(* IEC 61131-3 sources: HypervisionPLC-SCADA/demo/varme-plc, 5 files *)

(* ---- globals.st ---- *)
GLOBAL_VAR
  g_cmd    : INT;   (* L1: b0-3 P1-P4, b4 MVS1, b5 MVS2, b6 pille, b7 VP *)
  g_fb     : INT;   (* L2: b0-3 pumpe koerer, b6 pilleflamme, b9 FF-flamme, b10 Laddomat, b11 pillefejl *)
  g_fault  : INT;   (* L4: b0-3 pumpefejl, b4 pille, b5 laekage, b7 VP; b12 VP-fejlsignal *)
  g_speed  : REAL;  (* L4: tidsfaktor *)
  g_tude   : REAL;  (* L4: udetemp *)
  g_att1   : REAL;  (* L3: tank top *)
  g_att3   : REAL;  (* L3: tank midt *)
  g_att6   : REAL;  (* L3: tank bund *)
  g_fftf   : REAL;  (* L2 *)
  g_pftf   : REAL;  (* L2 *)
  g_mch    : REAL;  (* L2: ladeflow til tank kg/s *)
  g_tch    : REAL;  (* L2: ladetemp *)
  g_str    : REAL;  (* L3: vandet til M1 = pillefyrets indloeb (STR eller tanktop) *)
  g_vptf   : REAL;  (* L4: VP-fremloeb til tanken *)
  g_stf_sp : REAL;  (* L1: fremloebssetpunkt *)
  g_tryk   : REAL;  (* L4: bar *)
END_VAR

(* ---- logic1_styring.st ---- *)
PROGRAM Styring
(* Demo-varmeanlaeg, Logic1: styringen (det en rigtig PLC ville goere).
   Laeser anlaeggets tilstand fra GLOBAL_VAR og skriver kommandoer i g_cmd.
   cmd_mode: 0 Auto, 1 Manuel mode 1, 2 Manuel mode 2, 3 Manuel mode 3.
   MODE 1 Hus + pille (M1 AB-A, M2 AB-A, P1) - 2 Hus + pille + tank (M1 AB-A, M2 AB-B, P1)
   - 3 Hus + tank (M1 AB-B, M2 AB-B, P2). Auto: tanken ind (mode 3) ved ATT1 >= sp_tank_ind,
   ud (mode 1) under sp_tank_ud. Varmepumpen startes manuelt (cmd_vp). Interval 500 ms. *)
VAR
  SMS_TXT      : STRING;
  cmd_mode     : INT;
  cmd_kvitter  : BOOL;
  cmd_vp       : BOOL;
  sp_rum       : REAL := 21.0;
  sp_kurve     : REAL := 1.0;
  sp_stf_max   : REAL := 55.0;
  sp_tank_ind  : REAL := 60.0;
  sp_tank_ud   : REAL := 45.0;
  sp_vp_min    : REAL;          (* -5,0 saettes ved foerste scan: negative startvaerdier bliver 0 i firmwaren *)
  MODE         : INT := 1;
  SMS          : INT;
  STF_SP       : REAL;
  TANK_IND     : BOOL;
  PS1          : BOOL;
  PS2          : BOOL;
  PS3          : BOOL;
  PS4          : BOOL;
  F_HUS        : BOOL;
  F_PILLE      : BOOL;
  F_TANK       : BOOL;
  F_BYPASS     : BOOL;
  AL_P1        : BOOL;
  AL_P2        : BOOL;
  AL_P3        : BOOL;
  AL_P4        : BOOL;
  AL_VP        : BOOL;
  AL_PILLE     : BOOL;
  AL_TRYK_LAV  : BOOL;
  AL_TRYK_HOEJ : BOOL;
  AL_FF_TEMP   : BOOL;
  AL_TANK_KOLD : BOOL;
  ALARMER      : INT;
  kv           : BOOL;
  fb           : INT;
  cmd          : INT;
  tude         : REAL;
  t1           : REAL;
  trykstop     : BOOL;
  c_p1         : BOOL;
  c_p2         : BOOL;
  c_p3         : BOOL;
  c_p4         : BOOL;
  c_pille      : BOOL;
  c_vp         : BOOL;
  init         : BOOL;
END_VAR
BEGIN
  IF NOT init THEN sp_vp_min := -5.0; init := TRUE; END_IF;
  kv := cmd_kvitter;
  cmd_kvitter := FALSE;
  fb := g_fb;
  tude := g_tude;
  t1 := g_att1;

  (* Pumpefejl: kommanderet, men ingen tilbagemelding i 10 s -> laast til kvittering *)
  AL_P1 := SR(TON(BIT_TST(g_cmd, 0) AND NOT BIT_TST(fb, 0), T#10s), kv);
  AL_P2 := SR(TON(BIT_TST(g_cmd, 1) AND NOT BIT_TST(fb, 1), T#10s), kv);
  AL_P3 := SR(TON(BIT_TST(g_cmd, 2) AND NOT BIT_TST(fb, 2), T#10s), kv);
  AL_P4 := SR(TON(BIT_TST(g_cmd, 3) AND NOT BIT_TST(fb, 3), T#10s), kv);
  AL_VP := SR(BIT_TST(g_fault, 12), kv);   (* fejlsignal fra VP'ens egen styring *)
  AL_PILLE := SR(BIT_TST(fb, 11), kv);
  AL_TRYK_LAV := g_tryk < 1.0;
  AL_TRYK_HOEJ := g_tryk > 2.4;
  AL_FF_TEMP := g_fftf > 95.0;
  trykstop := g_tryk < 0.6;

  STF_SP := LIMIT(20.0, sp_rum + sp_kurve * (sp_rum - tude), sp_stf_max);
  g_stf_sp := STF_SP;

  (* Tanken i kredsen (Auto): ind ved sp_tank_ind, ud under sp_tank_ud *)
  IF t1 >= sp_tank_ind THEN
    TANK_IND := TRUE;
  ELSIF t1 < sp_tank_ud THEN
    TANK_IND := FALSE;
  END_IF;
  IF cmd_mode = 0 THEN
    IF TANK_IND THEN MODE := 3; ELSE MODE := 1; END_IF;
  ELSE
    MODE := LIMIT(1, cmd_mode, 3);
  END_IF;
  AL_TANK_KOLD := (cmd_mode = 3) AND (t1 < STF_SP - 5.0);

  c_p1 := MODE < 3;                 (* P1 i pillefyrets sloejfe: mode 1 og 2 *)
  c_p2 := MODE = 3;                 (* P2 fra tanken: mode 3 *)
  c_pille := c_p1 AND NOT AL_PILLE;
  c_vp := cmd_vp AND (tude >= sp_vp_min) AND NOT AL_VP AND NOT AL_P3;
  c_p3 := c_vp;
  c_p4 := HYSTERESIS(g_fftf, 60.0, 55.0);   (* Laddomat-pumpen koerer altid naar braendefyret er varmt *)

  SMS := MODE;
  IF trykstop THEN
    c_p1 := FALSE; c_p2 := FALSE; c_p3 := FALSE; c_pille := FALSE; c_vp := FALSE;
    SMS := 10;
  END_IF;
  c_p1 := c_p1 AND NOT AL_P1;
  c_p2 := c_p2 AND NOT AL_P2;
  c_p3 := c_p3 AND NOT AL_P3;
  c_p4 := c_p4 AND NOT AL_P4;
  c_vp := c_vp AND c_p3;

  cmd := 0;
  IF c_p1 THEN cmd := BIT_SET(cmd, 0); END_IF;
  IF c_p2 THEN cmd := BIT_SET(cmd, 1); END_IF;
  IF c_p3 THEN cmd := BIT_SET(cmd, 2); END_IF;
  IF c_p4 THEN cmd := BIT_SET(cmd, 3); END_IF;
  IF MODE = 3 THEN cmd := BIT_SET(cmd, 4); END_IF;    (* MVS1 AB-B *)
  IF MODE >= 2 THEN cmd := BIT_SET(cmd, 5); END_IF;   (* MVS2 AB-B *)
  IF c_pille THEN cmd := BIT_SET(cmd, 6); END_IF;
  IF c_vp THEN cmd := BIT_SET(cmd, 7); END_IF;
  g_cmd := cmd;

  (* SMS: 1-3 mode, 10 trykstop *)
  CASE SMS OF
    1: SMS_TXT := 'Hus + pille';
    2: SMS_TXT := 'Hus + pille + tank';
    3: SMS_TXT := 'Hus + tank';
    10: SMS_TXT := 'TRYKSTOP';
  END_CASE;
  PS1 := BIT_TST(fb, 0);
  PS2 := BIT_TST(fb, 1);
  PS3 := BIT_TST(fb, 2);
  PS4 := BIT_TST(fb, 3);
  (* Kredsdele med flow (roerene paa tegningen) *)
  F_HUS := PS1 OR PS2;
  F_PILLE := PS1;
  F_TANK := F_HUS AND (MODE >= 2);
  F_BYPASS := PS1 AND (MODE = 1);
  ALARMER := BOOL_TO_INT(AL_P1) + BOOL_TO_INT(AL_P2) + BOOL_TO_INT(AL_P3) + BOOL_TO_INT(AL_P4)
           + BOOL_TO_INT(AL_VP) + BOOL_TO_INT(AL_PILLE) + BOOL_TO_INT(AL_TRYK_LAV)
           + BOOL_TO_INT(AL_TRYK_HOEJ) + BOOL_TO_INT(AL_FF_TEMP) + BOOL_TO_INT(AL_TANK_KOLD);
END_PROGRAM

(* ---- logic2_kilder.st ---- *)
PROGRAM Kilder
(* Demo-varmeanlaeg, Logic2: procesmodel for braendefyr (+ Laddomat/P4) og
   pillefyr (i husets kreds med P1, mode 1 og 2); varmepumpen og braendefyrets statustekst ligger i Logic4.
   Leverer braendefyrets ladeflow/-temp til tanken (g_mch/g_tch) og tilbagemeldinger i g_fb.
   Pillefyrets indloeb: g_str (vandet til M1, fra Logic3). Interval 500 ms. *)
VAR
  PILLE_TXT  : STRING;
  cmd_fyr_op : BOOL;
  sp_pille   : REAL := 75.0;
  FFTF       : REAL := 20.0;
  FFTR       : REAL := 20.0;
  FF_KW      : REAL;
  FF_KG      : REAL;
  LADDOMAT   : BOOL;
  PFTF       : REAL := 20.0;
  PFTR       : REAL := 20.0;
  PILLE_KW   : REAL;
  PILLE_KG   : REAL;
  PILLE_ST   : INT;
  PILLE_STARTS : DINT;
  E_FF       : REAL;
  E_PILLE    : REAL;
  dt         : REAL;
  cmd        : INT;
  flt        : INT;
  fb         : INT;
  r_p1       : BOOL;
  r_p2       : BOOL;
  r_p4       : BOOL;
  ff_q       : REAL;
  ff_mt      : REAL;
  psp        : REAL;
  ps_t       : REAL;
  p_q        : REAL;
  pm         : REAL;
  pret       : REAL;
  en         : BOOL;
END_VAR
BEGIN
  dt := 0.5 * MAX(g_speed, 1.0);
  cmd := g_cmd;
  flt := g_fault;
  (* pumper der faktisk koerer: kommanderet og ikke i fejl *)
  r_p1 := BIT_TST(cmd, 0) AND NOT BIT_TST(flt, 0);
  r_p2 := BIT_TST(cmd, 1) AND NOT BIT_TST(flt, 1);
  r_p4 := BIT_TST(cmd, 3) AND NOT BIT_TST(flt, 3);
  fb := 0;
  IF r_p1 THEN fb := BIT_SET(fb, 0); END_IF;
  IF r_p2 THEN fb := BIT_SET(fb, 1); END_IF;
  IF BIT_TST(cmd, 2) AND NOT BIT_TST(flt, 2) THEN fb := BIT_SET(fb, 2); END_IF;
  IF r_p4 THEN fb := BIT_SET(fb, 3); END_IF;

  (* ---- Braendefyr: 15 kg pr. ilaegning, maks 30 kg, 25 kW, spjaeld over 88 C ---- *)
  IF cmd_fyr_op THEN FF_KG := MIN(FF_KG + 15.0, 30.0); END_IF;
  cmd_fyr_op := FALSE;
  IF FF_KG > 0.0 THEN
    FF_KW := 25.0 * MIN(1.0, FF_KG / 4.0) * LIMIT(0.3, (FFTF - 10.0) / 50.0, 1.0);
    IF FFTF > 88.0 THEN FF_KW := FF_KW * 0.3; END_IF;
  ELSE
    FF_KW := 0.0;
  END_IF;
  FF_KG := FF_KG - FF_KW * dt / 12000.0;
  IF FF_KG < 0.3 THEN FF_KG := 0.0; END_IF;   (* gloederne er braendt ud *)
  LADDOMAT := HYSTERESIS(FFTF, 72.0, 68.0);
  ff_q := 0.0; ff_mt := 0.0;
  IF r_p4 THEN
    IF LADDOMAT THEN
      FFTR := MIN(MAX(g_att6, 60.0), FFTF);
      ff_q := 0.3 * 4.186 * (FFTF - FFTR);
      ff_mt := ff_q / (4.186 * MAX(FFTF - g_att6, 2.0));
    ELSE
      FFTR := FFTF - 1.0;
    END_IF;
  ELSE
    FFTR := FFTR + (20.0 - FFTR) * MIN(1.0, dt / 1800.0);
  END_IF;
  FFTF := LIMIT(0.0, FFTF + (FF_KW - ff_q - 0.05 * (FFTF - 20.0)) * dt / 400.0, 112.0);
  g_fftf := FFTF;
  E_FF := E_FF + ff_q * dt / 3600.0;

  (* ---- Pillefyr: 0 Stop, 1 Taending, 2 Drift (5-15 kW), 3 Udbraending, 4 Fejl ---- *)
  en := BIT_TST(cmd, 6);
  psp := MIN(sp_pille, g_stf_sp + 5.0);   (* varmer husets vand direkte *)
  CASE PILLE_ST OF
    0: PILLE_KW := 0.0;
       IF en AND (PFTF < psp - 5.0) THEN PILLE_ST := 1; ps_t := 0.0; PILLE_STARTS := PILLE_STARTS + 1; END_IF;
    1: PILLE_KW := 0.5;
       ps_t := ps_t + dt;
       IF NOT en THEN PILLE_ST := 0;
       ELSIF BIT_TST(flt, 4) THEN
         IF ps_t > 600.0 THEN PILLE_ST := 4; END_IF;
       ELSIF ps_t > 180.0 THEN PILLE_ST := 2;
       END_IF;
    2: PILLE_KW := LIMIT(5.0, 5.0 + (psp - PFTF) * 1.5, 15.0);
       IF (NOT en) OR (PFTF > psp + 5.0) THEN PILLE_ST := 3; ps_t := 0.0; END_IF;
    3: ps_t := ps_t + dt;
       PILLE_KW := MAX(0.0, 3.0 - ps_t * 0.01);
       IF ps_t > 300.0 THEN PILLE_ST := 0; END_IF;
    4: PILLE_KW := 0.0;
       IF NOT en THEN PILLE_ST := 0; END_IF;
  END_CASE;
  pm := 0.0; pret := PFTR;
  IF r_p1 THEN pm := 0.25; pret := g_str; END_IF;   (* P1: 15 L/min gennem pillefyret *)
  IF pm > 0.0 THEN
    PFTR := pret;
  ELSE
    PFTR := PFTR + (20.0 - PFTR) * MIN(1.0, dt / 1800.0);
  END_IF;
  p_q := pm * 4.186 * (PFTF - pret);
  PFTF := LIMIT(0.0, PFTF + (PILLE_KW - p_q - 0.03 * (PFTF - 20.0)) * dt / 250.0, 112.0);
  g_pftf := PFTF;
  E_PILLE := E_PILLE + MAX(p_q, 0.0) * dt / 3600.0;
  PILLE_KG := PILLE_KG + PILLE_KW * dt / 15552.0;
  CASE PILLE_ST OF
    0: PILLE_TXT := 'Stop';
    1: PILLE_TXT := 'Tænding';
    2: PILLE_TXT := 'Drift';
    3: PILLE_TXT := 'Udbrænding';
    4: PILLE_TXT := 'Fejl';
  END_CASE;

  (* ---- Ladning af tanken fra braendefyret (Laddomat) ---- *)
  g_mch := ff_mt;
  g_tch := FFTF;

  IF PILLE_ST = 2 THEN fb := BIT_SET(fb, 6); END_IF;
  IF FF_KG > 0.0 THEN fb := BIT_SET(fb, 9); END_IF;
  IF LADDOMAT THEN fb := BIT_SET(fb, 10); END_IF;
  IF PILLE_ST = 4 THEN fb := BIT_SET(fb, 11); END_IF;
  g_fb := fb;
END_PROGRAM

(* ---- logic3_tank_hus.st ---- *)
PROGRAM TankHus
(* Demo-varmeanlaeg, Logic3: akkumuleringstank i 6 lag (750 L), husets
   varmekreds med AVTB-blandeventil og P1, motorventiler MVS1/MVS2
   (30 s gangtid i realtid). Interval 500 ms. *)
VAR
  MVS1_TXT : STRING;
  MVS2_TXT : STRING;
  T        : ARRAY[1..6] OF REAL;
  ATT1     : REAL;
  ATT2     : REAL;
  ATT3     : REAL;
  ATT4     : REAL;
  ATT5     : REAL;
  ATT6     : REAL;
  ATF      : REAL;
  TS       : REAL;
  E_TANK   : REAL;
  STF      : REAL := 30.0;
  STR      : REAL := 30.0;
  MVT2     : REAL := 30.0;
  FMTR     : REAL;
  T_RUM    : REAL := 21.0;
  Q_HUS    : REAL;
  E_HUS    : REAL;
  MVS1_POS : REAL;
  MVS2_POS : REAL;
  cmd_mvs1 : INT;
  cmd_mvs2 : INT;
  init     : BOOL;
  w        : BOOL;
  i        : INT;
  dt       : REAL;
  k        : REAL;
  m_h      : REAL;
  m_ht     : REAL;
  m_ch     : REAL;
  net      : REAL;
  up       : REAL;
  down     : REAL;
  prev     : REAL;
  old      : REAL;
  avg      : REAL;
  frac     : REAL;
  tsrc     : REAL;
  sum      : REAL;
  tch      : REAL;
  tin      : REAL;
END_VAR
BEGIN
  IF NOT init THEN
    FOR i := 1 TO 6 DO T[i] := 52.0 - 3.0 * INT_TO_REAL(i); END_FOR;
    init := TRUE;
  END_IF;
  dt := 0.5 * MAX(g_speed, 1.0);

  (* Motorventiler: ON = AB-B, OFF = AB-A. MVS1 AB-B = P2-grenen (uden om pillefyret), MVS2 AB-B = tanken i kredsen *)
  (* Haandbetjening paa motoren: cmd_mvsN 0 = Auto (styringen), 1 = AB-A, 2 = AB-B *)
  w := BIT_TST(g_cmd, 4);
  IF cmd_mvs1 = 1 THEN w := FALSE; ELSIF cmd_mvs1 = 2 THEN w := TRUE; END_IF;
  IF w THEN MVS1_POS := MIN(100.0, MVS1_POS + 1.667); ELSE MVS1_POS := MAX(0.0, MVS1_POS - 1.667); END_IF;
  w := BIT_TST(g_cmd, 5);
  IF cmd_mvs2 = 1 THEN w := FALSE; ELSIF cmd_mvs2 = 2 THEN w := TRUE; END_IF;
  IF w THEN MVS2_POS := MIN(100.0, MVS2_POS + 1.667); ELSE MVS2_POS := MAX(0.0, MVS2_POS - 1.667); END_IF;
  IF MVS1_POS >= 100.0 THEN MVS1_TXT := 'AB-B'; ELSIF MVS1_POS <= 0.0 THEN MVS1_TXT := 'AB-A'; ELSE MVS1_TXT := 'Kører'; END_IF;
  IF MVS2_POS >= 100.0 THEN MVS2_TXT := 'AB-B'; ELSIF MVS2_POS <= 0.0 THEN MVS2_TXT := 'AB-A'; ELSE MVS2_TXT := 'Kører'; END_IF;

  (* Husets kreds: P1 eller P2 = 15 L/min. M2: retur direkte (AB-A) eller gennem tanken (AB-B);
     M1: gennem pillefyret (AB-A) eller uden om (AB-B). AVTB blander ned til fremloebssetpunktet *)
  m_h := 0.0;
  IF BIT_TST(g_fb, 0) OR BIT_TST(g_fb, 1) THEN m_h := 0.25; END_IF;
  tin := SEL(MVS2_POS > 50.0, STR, T[1]);
  g_str := tin;   (* pillefyrets indloeb *)
  tsrc := SEL(MVS1_POS > 50.0, g_pftf, tin);
  frac := 1.0;
  IF tsrc > STR + 0.5 THEN frac := LIMIT(0.0, (g_stf_sp - STR) / (tsrc - STR), 1.0); END_IF;
  IF m_h > 0.0 THEN
    STF := STR + frac * (tsrc - STR);
    Q_HUS := MAX(0.0, 0.285 * (STF - T_RUM) / (1.0 + 0.285 / (2.0 * m_h * 4.186)));
    STR := STF - Q_HUS / (m_h * 4.186);
  ELSE
    Q_HUS := 0.0;
    STF := STF + (T_RUM - STF) * MIN(1.0, dt / 1200.0);
    STR := STR + (T_RUM - STR) * MIN(1.0, dt / 1200.0);
  END_IF;
  T_RUM := T_RUM + (Q_HUS + 0.4 - 0.25 * (T_RUM - g_tude)) * dt / 15000.0;
  FMTR := m_h * 60.0;
  MVT2 := STR;
  E_HUS := E_HUS + Q_HUS * dt / 3600.0;
  m_ht := 0.0;
  IF MVS2_POS > 50.0 THEN m_ht := m_h * frac; END_IF;   (* gennem tanken: retur i bunden, ud i toppen *)

  (* Tank: ladning i toppen fra kilderne, husets retur i bunden, lagdelt strømning *)
  m_ch := g_mch;
  IF BIT_TST(g_fb, 2) THEN   (* varmepumpen (P3) lader fra bund til top *)
    m_ch := m_ch + 0.3;
    tch := (g_mch * g_tch + 0.3 * g_vptf) / m_ch;
  ELSE
    tch := g_tch;
  END_IF;
  net := m_ch - m_ht;
  down := MAX(net, 0.0);
  up := MAX(0.0 - net, 0.0);
  k := dt / 125.0;
  prev := T[1];
  T[1] := T[1] + (m_ch * (tch - T[1]) + up * (T[2] - T[1])) * k;
  FOR i := 2 TO 5 DO
    old := T[i];
    T[i] := T[i] + (down * (prev - T[i]) + up * (T[i + 1] - T[i])) * k;
    prev := old;
  END_FOR;
  T[6] := T[6] + (down * (prev - T[6]) + m_ht * (STR - T[6])) * k;
  sum := 0.0;
  FOR i := 1 TO 6 DO
    T[i] := T[i] - 0.002 * (T[i] - 20.0) * dt / 523.0;
    sum := sum + T[i];
  END_FOR;
  FOR i := 1 TO 5 DO
    IF T[i + 1] > T[i] THEN
      avg := (T[i] + T[i + 1]) / 2.0;
      T[i] := avg;
      T[i + 1] := avg;
    END_IF;
  END_FOR;

  ATT1 := T[1]; ATT2 := T[2]; ATT3 := T[3]; ATT4 := T[4]; ATT5 := T[5]; ATT6 := T[6];
  ATF := T[1];
  E_TANK := 0.14535 * (sum - 180.0);
  TS := LIMIT(0.0, (sum / 6.0 - 30.0) * 2.0, 100.0);
  g_att1 := T[1];
  g_att3 := T[3];
  g_att6 := T[6];
END_PROGRAM

(* ---- logic4_system.st ---- *)
PROGRAM SystemDemo
(* Demo-varmeanlaeg, Logic4: systemtryk med ekspansion og sikkerhedsventiler
   (2,5 bar), udetemperatur over doegnet, simuleret klokke, tidsfaktor,
   scenarier og fejlinjektion, samt varmepumpen (P3). Interval 500 ms.
   cmd_scenarie: 0 Normal, 1 Vinternat, 2 Sommer, 3 Laekage, 4 Pumpefejl P1. *)
VAR
  FFS_TXT       : STRING;   (* braendefyrets status *)
  sp_speed      : REAL := 1.0;
  cmd_scenarie  : INT;
  cmd_efterfyld : BOOL;
  sp_tude_fast  : BOOL;
  sp_tude       : REAL := 5.0;
  f_P1          : BOOL;
  f_P2          : BOOL;
  f_P3          : BOOL;
  f_P4          : BOOL;
  f_pille       : BOOL;
  f_vp          : BOOL;
  f_laek        : BOOL;
  ST            : REAL := 1.2;
  SV_AABEN      : BOOL;
  T_UDE         : REAL;
  KLOKKE        : REAL;
  DAG           : INT;
  p_fill        : REAL := 1.2;
  t_dag         : REAL := 21600.0;
  dt            : REAL;
  mid           : REAL;
  amp           : REAL;
  tm            : REAL;
  p             : REAL;
  flt           : INT;
  VPTF          : REAL := 20.0;
  VPTR          : REAL := 20.0;
  VP_KW         : REAL;
  VP_EL         : REAL;
  VP_COP        : REAL := 4.0;
  VP_RUN        : BOOL;
  E_VP          : REAL;
  E_VP_EL       : REAL;
  r_p3          : BOOL;
  vq            : REAL;
  kf            : REAL;
END_VAR
BEGIN
  sp_speed := LIMIT(1.0, sp_speed, 120.0);
  g_speed := sp_speed;
  dt := 0.5 * sp_speed;

  t_dag := t_dag + dt;
  IF t_dag >= 86400.0 THEN t_dag := t_dag - 86400.0; DAG := DAG + 1; END_IF;
  KLOKKE := t_dag / 3600.0;

  CASE cmd_scenarie OF
    1: mid := -12.0; amp := 3.0;
    2: mid := 18.0; amp := 6.0;
  ELSE
    mid := 3.0; amp := 4.0;
  END_CASE;
  (* koldest kl. 05, varmest kl. 17 *)
  T_UDE := mid - amp * COS((t_dag - 18000.0) * 0.0000727221);
  IF sp_tude_fast THEN T_UDE := sp_tude; END_IF;
  g_tude := T_UDE;

  flt := 0;
  IF f_P1 OR (cmd_scenarie = 4) THEN flt := BIT_SET(flt, 0); END_IF;
  IF f_P2 THEN flt := BIT_SET(flt, 1); END_IF;
  IF f_P3 THEN flt := BIT_SET(flt, 2); END_IF;
  IF f_P4 THEN flt := BIT_SET(flt, 3); END_IF;
  IF f_pille THEN flt := BIT_SET(flt, 4); END_IF;
  IF f_laek OR (cmd_scenarie = 3) THEN flt := BIT_SET(flt, 5); END_IF;
  IF f_vp THEN flt := BIT_SET(flt, 7); END_IF;

  (* ---- Varmepumpe: ca. 8 kW, COP efter udetemp og fremloeb, maks 65 C fremloeb, stopper ved retur >= 58 C ---- *)
  r_p3 := BIT_TST(g_cmd, 2) AND NOT f_P3;
  VP_RUN := BIT_TST(g_cmd, 7) AND r_p3 AND NOT f_vp AND (g_att6 < 58.0);
  IF BIT_TST(g_cmd, 7) AND f_vp THEN flt := BIT_SET(flt, 12); END_IF;
  g_fault := flt;
  vq := 0.0;
  IF VP_RUN THEN
    vq := 8.0 * (1.0 + 0.02 * (T_UDE - 7.0));
    VP_COP := LIMIT(1.5, 4.8 - 0.07 * (VPTF - 35.0) + 0.06 * (T_UDE - 7.0), 6.0);
  END_IF;
  kf := MIN(1.0, dt / 1800.0);
  VP_KW := VP_KW + (vq - VP_KW) * MIN(1.0, dt / 120.0);
  IF r_p3 THEN
    VPTR := g_att6;
    VPTF := MIN(65.0, g_att6 + VP_KW / 1.2558);
  ELSE
    VP_KW := 0.0;
    VPTF := VPTF + (20.0 - VPTF) * kf;
    VPTR := VPTR + (20.0 - VPTR) * kf;
  END_IF;
  g_vptf := VPTF;
  VP_EL := 0.0;
  IF VP_RUN THEN VP_EL := VP_KW / VP_COP; END_IF;
  E_VP := E_VP + VP_KW * dt / 3600.0;
  E_VP_EL := E_VP_EL + VP_EL * dt / 3600.0;

  (* Tryk: fyldning + varmeudvidelse (ekspansionsbeholder) + damp over 100 C *)
  tm := (g_att1 + g_att3 + g_att6) / 3.0 * 0.85 + (g_fftf + g_pftf) * 0.075;
  p := p_fill + 0.012 * (tm - 20.0);
  IF g_fftf > 100.0 THEN p := p + (g_fftf - 100.0) * 0.15; END_IF;
  IF g_pftf > 100.0 THEN p := p + (g_pftf - 100.0) * 0.15; END_IF;
  SV_AABEN := HYSTERESIS(p, 2.5, 2.3);
  IF SV_AABEN THEN p_fill := p_fill - 0.002 * dt; END_IF;
  IF BIT_TST(flt, 5) THEN p_fill := p_fill - 0.00005 * dt; END_IF;
  IF cmd_efterfyld THEN p_fill := 1.2; END_IF;
  cmd_efterfyld := FALSE;
  p_fill := MAX(p_fill, 0.0);
  ST := MAX(p, 0.0);
  g_tryk := ST;
  IF g_fftf > 95.0 THEN FFS_TXT := 'Overtemp';
  ELSIF BIT_TST(g_fb, 9) AND (g_fftf < 60.0) THEN FFS_TXT := 'Optænding';
  ELSIF BIT_TST(g_fb, 9) THEN FFS_TXT := 'Drift';
  ELSE FFS_TXT := 'Slukket';
  END_IF;
  WDT_FEED();
END_PROGRAM
